Fanuc KAREL source: KX00024.KL

PROGRAM KX00024
%NOLOCKGROUP
VAR
  I: INTEGER
  J: INTEGER
  B: BOOLEAN
  F: FILE
  S: STRING[80]
  P: XYZWPR
  CNF: CONFIG
BEGIN
  CNF.CFG_FLIP = TRUE
  B = CNF.CFG_FLIP
END KX00024
